(* IEC 61131-3 sources: STruCpp/tests/st-validation/programs, 4 files *)

(* ---- configuration.st ---- *)
PROGRAM ConfigTest
  VAR
    cycle_count : INT;
    running : BOOL;
  END_VAR

  cycle_count := cycle_count + 1;
  running := TRUE;
END_PROGRAM

(* ---- multi_program.st ---- *)
PROGRAM Adder
  VAR
    a : INT;
    b : INT;
    result : INT;
  END_VAR
  result := a + b;
END_PROGRAM

PROGRAM Doubler
  VAR
    input : INT;
    output : INT;
  END_VAR
  output := input * 2;
END_PROGRAM

(* ---- test_configuration.st ---- *)
TEST 'Program state increments on each call'
  VAR uut : ConfigTest; END_VAR
  uut();
  ASSERT_EQ(uut.cycle_count, 1);
  ASSERT_TRUE(uut.running);
  uut();
  ASSERT_EQ(uut.cycle_count, 2);
END_TEST

(* ---- test_multi_program.st ---- *)
TEST 'Adder computes sum'
  VAR uut : Adder; END_VAR
  uut.a := 15;
  uut.b := 25;
  uut();
  ASSERT_EQ(uut.result, 40);
END_TEST

TEST 'Doubler computes double'
  VAR uut : Doubler; END_VAR
  uut.input := 7;
  uut();
  ASSERT_EQ(uut.output, 14);
END_TEST

TEST 'Programs are independent'
  VAR add : Adder; dbl : Doubler; END_VAR
  add.a := 3;
  add.b := 4;
  add();
  dbl.input := add.result;
  dbl();
  ASSERT_EQ(add.result, 7);
  ASSERT_EQ(dbl.output, 14);
END_TEST
